(* IEC 61131-3 sources: guidance-for-physical-ai-production-designer-on-aws/source/plan2cell/examples/cell_2robot/plc/trust/head/src, 14 files *)

(* ---- E_CellError.st ---- *)
(*
 * E_CellError
 *
 * Fault codes of the cell (FB_Cell.eError), the robot drivers (FB_VassRobot.eError)
 * and the zone arbiter (FB_ZoneArbiter.eFault). ERR_NONE = no fault.
 *)

TYPE E_CellError :
(
    ERR_NONE                := 0,

    (* VASS bring-up and job handshake (FB_VassRobot) *)
    ERR_SAFETY_TIMEOUT      := 10,      (* SafeIn0.0 / SafeIn1.4 not reported *)
    ERR_DRIVES_TIMEOUT      := 11,      (* DrivesOn not reported *)
    ERR_EXT_TIMEOUT         := 12,      (* EXT mode not reported *)
    ERR_NOT_READY           := 13,      (* robot not Ready (or JobAck stuck) before a job *)
    ERR_ACK_TIMEOUT         := 14,      (* no JobAck after JobRequest *)
    ERR_ECHO_MISMATCH       := 15,      (* echoed job number <> requested job number *)
    ERR_START_TIMEOUT       := 16,      (* ProgRunning not reported after ProgStart *)
    ERR_ROBOT_STOPPED       := 17,      (* ProgRunning dropped without ProgFinished (T_STOP_DEBOUNCE) *)
    ERR_ROBOT_ERROR         := 18,      (* robot reports Error *)
    ERR_SAFETY_LOST         := 19,      (* safe status lost while up *)
    ERR_STOP_TIMEOUT        := 20,      (* robot still running after Stop + Cancel *)
    ERR_RESET_FAILED        := 21,      (* robot still in error after Reset *)
    ERR_DRIVES_LOST         := 22,      (* DrivesOn lost while up *)
    ERR_UNEXPECTED_RUN      := 23,      (* ProgRunning reported outside a job (off / bring-up / idle) *)

    (* zone protocol and supervision (FB_ZoneArbiter, FB_Cell) *)
    ERR_OP_WATCHDOG         := 30,      (* op took longer than aOps[].tLimit *)
    ERR_ZONE_WAIT_TIMEOUT   := 31,      (* zone wait past aOps[].tZoneDeadline since cycle start *)
    ERR_STEP_SEQUENCE       := 32,      (* op index did not advance by exactly +1, or 0 between two ops *)
    ERR_REQ_MISMATCH        := 33,      (* REQUEST <> mask of the reported op (debounced) *)
    ERR_TICKET_SKIPPED      := 34,      (* own ticket for another op, or zone consumed (debounced) *)
    ERR_PROGRAM_INCOMPLETE  := 35,      (* job done but last op index <> op count *)
    ERR_RELEASE_INVALID     := 36,      (* REQUEST dropped by a robot that is not running OK *)
    ERR_ROBOT_STALLED       := 37,      (* zone op without REQUEST and grant, or op index 0 too long *)
    ERR_UNEXPECTED_REQUEST  := 38,      (* holder raised bits it was not granted *)
    ERR_TICKETS_LEFT        := 39,      (* cycle done with unconsumed tickets *)
    ERR_HOME_FAILED         := 40,      (* blind homing did not reach the home pose *)
    ERR_HANDSHAKE           := 41,      (* op index changed while a grant was held (4-phase violated) *)
    ERR_ZONE_BYPASSED       := 42,      (* zone / permit op left without ever being granted *)

    (* operator *)
    ERR_OPERATOR_STOP       := 50       (* bStop *)
);
END_TYPE

(* ---- E_CellState.st ---- *)
(*
 * E_CellState
 *
 * States of the cell controller FB_Cell.
 *)

TYPE E_CellState :
(
    CS_INIT                 := 0,       (* robots off *)
    CS_BRINGUP              := 10,      (* all robots: SAFETY_ENABLE -> DRIVES_ON -> MODE_EXT -> IDLE *)
    CS_HOMING_SELECT        := 20,      (* pick robot(s) not at home *)
    CS_HOMING_RUN           := 21,      (* blind homing with HOME_FOLGE *)
    CS_READY                := 30,      (* all robots at home, waiting for start / auto-run *)
    CS_START_JOBS           := 40,      (* production Folge commanded on every active robot *)
    CS_RUNNING              := 50,      (* robots run autonomously, zones arbitrated *)
    CS_CYCLE_DONE           := 60,      (* pause T_CYCLE_PAUSE before the next cycle *)
    CS_ABORTING             := 80,      (* grants dropped, Stop + Cancel to every busy robot *)
    CS_RECOVERY             := 85,      (* after an abort mid-cycle, or a start-up with an active robot
                                           away from home: wait for bRecoveryConfirm *)
    CS_RESETTING            := 90,      (* Reset to robots in error (an operator stop cancels it) *)
    CS_ERROR                := 99       (* latched until bReset *)
);
END_TYPE

(* ---- E_GrantPolicy.st ---- *)
(*
 * E_GrantPolicy
 *
 * Zone grant policy of FB_ZoneArbiter (GVL_Cell.GRANT_POLICY).
 *)

TYPE E_GrantPolicy :
(
    GP_PLANNED  := 0,       (* zone granted only to its next ticket holder (BT order) *)
    GP_FCFS     := 1        (* oldest request first - BT order NOT enforced *)
);
END_TYPE

(* ---- E_RobotState.st ---- *)
(*
 * E_RobotState
 *
 * States of the VASS driver FB_VassRobot (one robot).
 *)

TYPE E_RobotState :
(
    RS_OFF                  := 0,       (* outputs off, waiting for bPowerOn *)
    RS_SAFETY_ENABLE        := 1,       (* SafeOut0/1 set, waiting for safe status *)
    RS_DRIVES_ON            := 2,       (* DrivesOn requested *)
    RS_MODE_EXT             := 3,       (* EXT mode requested *)
    RS_IDLE                 := 10,      (* up, no job *)
    RS_JOB_WAIT_READY       := 20,      (* waiting for Ready and no JobAck *)
    RS_JOB_SEND             := 21,      (* job number + JobRequest, waiting for JobAck *)
    RS_JOB_START            := 22,      (* ProgStart pulse *)
    RS_JOB_WAIT_RUNNING     := 23,      (* waiting for ProgRunning (or ProgFinished) *)
    RS_JOB_RUNNING          := 24,      (* program running *)
    RS_JOB_DONE             := 25,      (* ProgFinished seen, bJobDone set *)
    RS_STOPPING             := 30,      (* Stop + Cancel held *)
    RS_RESET                := 40,      (* Reset held *)
    RS_ERROR                := 99       (* latched until bCmdReset *)
);
END_TYPE

(* ---- ST_OpInfo.st ---- *)
(*
 * ST_OpInfo
 *
 * One op of one robot (GVL_Cell.aOps). Op k of robot r is
 * GVL_Cell.aOps[GVL_Cell.anRobotFirstOp[r] + k - 1].
 *)

TYPE ST_OpInfo :
STRUCT
    nRobot              : INT;      (* robot index, 1-based *)
    nOp                 : INT;      (* op index of that robot, 1-based *)
    dwZoneMask          : DWORD;    (* REQUEST/GRANT mask: zone bits 0..30, bit 31 = permit *)
    nPredFirst          : INT;      (* permit preds: GVL_Cell.aPreds[nPredFirst .. nPredFirst + nPredCount - 1] *)
    nPredCount          : INT;      (* 0 = no permit predecessors *)
    tExpected           : TIME;     (* nominal duration *)
    tLimit              : TIME;     (* op watchdog (from the grant, or from the step change if mask = 0) *)
    tZoneDeadline       : TIME;     (* latest grant time since cycle start *)
    sName               : STRING(32);
END_STRUCT
END_TYPE

(* ---- ST_RobotIn.st ---- *)
(*
 * ST_RobotIn
 *
 * Copy of one robot's input image (robot -> PLC), filled by PLC_PRG from
 * GVL_IO.bySafeIn0_<tag>..bySafeIn7_<tag> and GVL_IO.aVassInputData_<tag>.
 *)

TYPE ST_RobotIn :
STRUCT
    abySafeIn           : ARRAY[0..7] OF BYTE;      (* PROFIsafe FDIO64 safe status *)
    aVassIn             : ARRAY[0..31] OF BYTE;     (* VASS DIO256 status telegram *)
END_STRUCT
END_TYPE

(* ---- ST_RobotOut.st ---- *)
(*
 * ST_RobotOut
 *
 * One robot's output image (PLC -> robot), copied by PLC_PRG to
 * GVL_IO.bySafeOut0_<tag>..bySafeOut7_<tag> and GVL_IO.aVassOutputData_<tag>.
 *)

TYPE ST_RobotOut :
STRUCT
    abySafeOut          : ARRAY[0..7] OF BYTE;      (* PROFIsafe FDIO64 safe commands *)
    aVassOut            : ARRAY[0..31] OF BYTE;     (* VASS DIO256 command telegram *)
END_STRUCT
END_TYPE

(* ---- ST_Ticket.st ---- *)
(*
 * ST_Ticket
 *
 * One (robot, op) reference: a zone ticket in GVL_Cell.aTickets or a permit
 * predecessor in GVL_Cell.aPreds. Both indices are 1-based; 0 = none (dummy row).
 *)

TYPE ST_Ticket :
STRUCT
    nRobot              : INT;      (* robot index 1..GVL_Cell.N_ROBOTS *)
    nOp                 : INT;      (* op index of that robot 1..anRobotOpCount[nRobot] *)
END_STRUCT
END_TYPE

(* ---- GVL_Cell.st ---- *)
NAMESPACE GVL_Cell
(*
 * GVL_Cell - generated by bt2plc 0.1.0 - DO NOT EDIT
 * Plan   : bt_1791274820_cell_2robot (cell cell_2robot)
 * Grants : planned ticket order
 *)
{attribute 'qualified_only'}
VAR_GLOBAL
    (* ========================================================================
       DIMENSIONS (array bounds are literals; *_DIM >= 1)
       ======================================================================== *)
    N_ROBOTS                : INT := 1;
    N_ZONES                 : INT := 0;
    N_OPS                   : INT := 2;
    N_PREDS                 : INT := 0;

    (* ========================================================================
       PROTOCOL / TIMING
       ======================================================================== *)
    PLAN_ID                 : WORD := WORD#16#A312;             (* fold of the plan fingerprint *)
    PROD_FOLGE              : WORD := WORD#11;                  (* default production Folge *)
    HOME_FOLGE              : WORD := WORD#125;                 (* blind homing *)
    JOB_NUMBER_BYTE         : BOOL := FALSE;                    (* FALSE: WORD LE bytes 2-3, TRUE: byte 2 *)
    PROFILE_VW              : BOOL := FALSE;                    (* TRUE: VW KS24 signal map and Folge handshake instead of the simulator telegram *)
    GRANT_POLICY            : E_GrantPolicy := E_GrantPolicy#GP_PLANNED;
    HOME_SEQUENTIAL         : BOOL := TRUE;
    AUTO_RUN                : BOOL := TRUE;                     (* start the next cycle automatically *)
    STEP_BYTE               : INT := 4;                         (* robot -> PLC, WORD LE op index *)
    REQ_BYTE                : INT := 28;                        (* robot -> PLC, DWORD LE zone requests *)
    GRANT_BYTE              : INT := 12;                        (* PLC -> robot, DWORD LE zone grants *)
    PLAN_ID_BYTE            : INT := 4;                         (* PLC -> robot, WORD LE plan id *)
    PERMIT_MASK             : DWORD := DWORD#16#80000000;       (* bit 31: permit predecessors *)
    T_RESET_PULSE           : TIME := T#1S;
    T_START_PULSE           : TIME := T#500MS;
    T_STOP_PULSE            : TIME := T#1S;
    T_HANDSHAKE             : TIME := T#5S;
    T_BRINGUP_LIMIT         : TIME := T#1M;                     (* safety enable: PROFINET connection set-up *)
    T_MISMATCH_DEBOUNCE     : TIME := T#200MS;
    T_STOP_DEBOUNCE         : TIME := T#200MS;                  (* job running: ProgRunning and ProgFinished low this long = robot stopped *)
    T_CYCLE_PAUSE           : TIME := T#2S;
    T_START_LIMIT           : TIME := T#15S;
    T_ABORT_LIMIT           : TIME := T#10S;
    T_HOME_LIMIT            : TIME := T#15S500MS;

    (* ========================================================================
       VW KS24 SIGNAL INDICES (used when PROFILE_VW; $IN/$OUT index, 1-based)
       ======================================================================== *)
    VW_READY_OUT            : INT := 9;                         (* O_R_Bereit *)
    VW_RK100_OUT            : INT := 10;                        (* O_R_RK100 safety circuit *)
    VW_AUTO_OUT             : INT := 12;                        (* O_R_Auto *)
    VW_ESTOP_OUT            : INT := 13;                        (* O_R_Notaus *)
    VW_END_OUT              : INT := 14;                        (* O_R_F_ENDE / LPKT *)
    VW_PF0_OUT              : INT := 15;                        (* O_R_PFO home position *)
    VW_STEP_OUT             : INT := 97;                        (* P_PktNr_SPS op index (16 bits) *)
    VW_REL_OUT              : INT := 41;                        (* interlock releases A41-56 *)
    VW_REQ_OUT              : INT := 81;                        (* interlock requests A81-96 *)
    VW_ERR_OUT              : INT := 225;                       (* VW_FEH_BIN_A error code (8 bits) *)
    VW_DRIVES_IN            : INT := 10;                        (* I_R_Ant_Ein *)
    VW_SRB_IN               : INT := 9;                         (* I_R_SRB Folge start *)
    VW_RESET_IN             : INT := 26;                        (* I_R_Quit_St acknowledge *)
    anInterlock             : ARRAY[1..1] OF INT := [0];        (* robot r, zone z -> VW interlock 1..16 (0 = not a member): index (r-1)*1+z *)

    (* ========================================================================
       ROBOTS (index = BT order)
       ======================================================================== *)
    asRobotTag              : ARRAY[1..1] OF STRING(16) := ['R1'];
    asRobotNs               : ARRAY[1..1] OF STRING(32) := ['robot1'];
    abRobotActive           : ARRAY[1..1] OF BOOL := [TRUE];
    abSafetyBypass          : ARRAY[1..1] OF BOOL := [FALSE];   (* SIMULATION ONLY: PROFIsafe slot-1 bits not required ([[robot]] safety_bypass) *)
    awRobotProdFolge        : ARRAY[1..1] OF WORD := [WORD#11];
    anRobotFirstOp          : ARRAY[1..1] OF INT := [1];        (* op k of robot r: aOps[anRobotFirstOp[r] + k - 1] *)
    anRobotOpCount          : ARRAY[1..1] OF INT := [2];

    (* ========================================================================
       ZONES - tickets of zone z: aTickets[anZoneFirst[z] .. anZoneFirst[z] + anZoneCount[z] - 1]
       ======================================================================== *)
    asZoneName              : ARRAY[1..1] OF STRING(8) := [''];
    anZoneFirst             : ARRAY[1..1] OF INT := [0];
    anZoneCount             : ARRAY[1..1] OF INT := [0];
    aTickets                : ARRAY[1..1] OF ST_Ticket := [
        (nRobot := 0, nOp := 0)    (* no zones *)
    ];

    (* ========================================================================
       OPS - op k of robot r: aOps[anRobotFirstOp[r] + k - 1]
       ======================================================================== *)
    (* tLimit = 1.5 x tExpected + 5 s ; tZoneDeadline = 1.5 x ASAP grant + (5 + 0.2) s x depth + 10 s *)
    aOps                    : ARRAY[1..2] OF ST_OpInfo := [
        (nRobot := 1, nOp := 1, dwZoneMask := DWORD#16#00000000, nPredFirst := 0, nPredCount := 0, tExpected := T#3S729MS, tLimit := T#10S594MS, tZoneDeadline := T#10S, sName := 'STAGE_R1'),    (* R1 #1 STAGE_R1 *)
        (nRobot := 1, nOp := 2, dwZoneMask := DWORD#16#00000000, nPredFirst := 0, nPredCount := 0, tExpected := T#2S419MS, tLimit := T#8S629MS, tZoneDeadline := T#20S794MS, sName := 'HOME')    (* R1 #2 HOME *)
    ];

    (* ========================================================================
       PERMIT PREDECESSORS - op preds: aPreds[nPredFirst .. nPredFirst + nPredCount - 1]
       ======================================================================== *)
    aPreds                  : ARRAY[1..1] OF ST_Ticket := [
        (nRobot := 0, nOp := 0)    (* no permit predecessors *)
    ];
END_VAR
END_NAMESPACE

(* ---- GVL_IO.st ---- *)
NAMESPACE GVL_IO
(*
 * GVL_IO - Head PLC I/O, one block per robot
 * Generated by bt2plc 0.1.0 for cell cell_2robot (plan bt_1791274820_cell_2robot)
 *
 * This is the PROFINET Controller (master) side.
 * From the controller's perspective:
 *   "Inputs"  = data received FROM the robot device (robot status)
 *   "Outputs" = data sent TO the robot device (PLC commands)
 *
 * Map in the I/O Mapping tab of each KUKA device under the PN-Controller:
 *   SafeIO_FDIO64_<tag> inputs  -> bySafeIn0_<tag>..bySafeIn7_<tag>
 *   SafeIO_FDIO64_<tag> outputs -> bySafeOut0_<tag>..bySafeOut7_<tag>
 *   VASS_DIO256_<tag> inputs    -> aVassInputData_<tag>
 *   VASS_DIO256_<tag> outputs   -> aVassOutputData_<tag>
 *
 * Only PLC_PRG accesses this GVL: whole arrays and single bytes are copied
 * into / out of FB_Cell (never write single elements of these arrays).
 *)

{attribute 'qualified_only'}
VAR_GLOBAL

    (* ========================================================================
       R1 - robot1 - kuka_robi1 (kuka-robi1, 192.168.100.11)
       ======================================================================== *)

    (* SLOT 1 - PROFIsafe FDIO64: safe status FROM robot (8 bytes) *)
    bySafeIn0_R1            : BYTE;     (* Byte 0: Drives OK, Stopped, Reduced speed... *)
    bySafeIn1_R1            : BYTE;     (* Byte 1: Gates, E-Stop, Enabling... *)
    bySafeIn2_R1            : BYTE;     (* Byte 2: STO, SS1, SS2, SOS, SLS... *)
    bySafeIn3_R1            : BYTE;
    bySafeIn4_R1            : BYTE;
    bySafeIn5_R1            : BYTE;
    bySafeIn6_R1            : BYTE;
    bySafeIn7_R1            : BYTE;

    (* SLOT 1 - PROFIsafe FDIO64: safe commands TO robot (8 bytes) *)
    bySafeOut0_R1           : BYTE;     (* Byte 0: Drive enable, E-Stop, SS1, SS2, SLS... *)
    bySafeOut1_R1           : BYTE;     (* Byte 1: Zone enables *)
    bySafeOut2_R1           : BYTE;
    bySafeOut3_R1           : BYTE;
    bySafeOut4_R1           : BYTE;
    bySafeOut5_R1           : BYTE;
    bySafeOut6_R1           : BYTE;
    bySafeOut7_R1           : BYTE;

    (* SLOT 2 - DIO256 VASS telegram (32 bytes each direction) *)
    aVassInputData_R1       : ARRAY[0..31] OF BYTE;         (* VASS status FROM robot *)
    aVassOutputData_R1      : ARRAY[0..31] OF BYTE;         (* VASS commands TO robot *)

END_VAR
END_NAMESPACE

(* ---- FB_Cell.st ---- *)
(*
 * FB_Cell
 * Generated by bt2plc 0.1.0 for cell cell_2robot (plan bt_1791274820_cell_2robot)
 *
 * Cell control for 1 robot(s): bring-up, blind homing (HOME_FOLGE), production
 * cycle (awRobotProdFolge started on every active robot; the robots run autonomously),
 * zone / permit arbitration (FB_ZoneArbiter), supervision (op index sequence, per-op
 * watchdog, zone-wait deadline, stall, program completeness), abort (stop all, drop grants,
 * rewind tickets), recovery confirmation and reset (Reset held >= 500 ms).
 *
 *   INIT -> BRINGUP -> HOMING_SELECT <-> HOMING_RUN -> READY -> START_JOBS -> RUNNING
 *        -> CYCLE_DONE -> READY ...
 *   any fault -> ABORTING -> ERROR -(bReset)-> RESETTING -> BRINGUP -> HOMING_SELECT ...
 *   abort with a robot inside its program (op index > 0, grant held, program left
 *   incomplete or away from home), or the first bring-up after INIT (head restart /
 *   download) with an active robot away from home:
 *        ... BRINGUP -> RECOVERY -(bRecoveryConfirm)-> RESETTING -> BRINGUP -> HOMING_SELECT
 *        (operator moves the robots clear in T1 first; homing is then always sequential)
 *   Start-up homing stays automatic when every active robot is at home.
 *
 * Operator: a bStop edge is latched in every state until it is consumed - abort (normal
 * states), cancel of the reset -> ERROR (INIT / RESETTING, driver Reset low), or cleared
 * (ERROR). A bReset edge in ABORTING is applied when ERROR is reached.
 *
 * Scan order: robot drivers (commands of the previous scan) -> op index tracking ->
 * faults known so far -> arbiter (this scan's inputs, no new grants after a fault) ->
 * watchdogs -> faults -> state machine -> GRANT bytes (0 when a fault is latched).
 * Op supervision runs whenever a robot's production job is commanded / running, in any
 * cell state: op index sequence, zone ops left without grant, op index 0 while running.
 *
 * Portable: one FB_VassRobot instance per robot (no FB instance arrays), timers are
 * TIME stamps of one free-running clock (_tNow).
 *)

FUNCTION_BLOCK FB_Cell
VAR_INPUT
    bEnable             : BOOL := TRUE;
    bAutoRun            : BOOL := TRUE;     (* Level: start a cycle whenever READY *)
    bStart              : BOOL;             (* Rising edge: start one cycle *)
    bStop               : BOOL;             (* Rising edge: abort (ERR_OPERATOR_STOP) *)
    bReset              : BOOL;             (* Rising edge in CS_ERROR: reset robots and cell *)
    bRecoveryConfirm    : BOOL;             (* Rising edge (from CS_ERROR on, while bRecoveryRequired): robots cleared *)
    astIn               : ARRAY[1..1] OF ST_RobotIn;    (* Robot inputs (copied from GVL_IO) *)
END_VAR

VAR_OUTPUT
    astOut              : ARRAY[1..1] OF ST_RobotOut;   (* Robot outputs (copied to GVL_IO) *)
    eState              : E_CellState;
    eError              : E_CellError;      (* First fault, ERR_NONE when OK *)
    nErrorRobot         : INT;              (* Robot of the fault, 0 = cell *)
    nErrorOp            : INT;              (* Op index of the fault, 0 = none *)
    nErrorZone          : INT;              (* Zone of the fault, 0 = none *)
    bCycleActive        : BOOL;             (* START_JOBS or RUNNING *)
    bError              : BOOL;             (* Fault latched until the reset is done *)
    bHomingRequired     : BOOL;         (* Profile vw-ks24: a robot is not at home and must be
                                           jogged there by the operator (no blind HOME Folge) *)
    bRecoveryRequired   : BOOL;             (* bRecoveryConfirm needed before homing (abort mid-cycle / start-up away from home) *)
    udiCycles           : UDINT;            (* Completed production cycles *)
    tLastCycle          : TIME;             (* Duration of the last cycle (RUNNING) *)
    aeRobotState        : ARRAY[1..1] OF E_RobotState;
    aeRobotError        : ARRAY[1..1] OF E_CellError;
    awStep              : ARRAY[1..1] OF WORD;          (* Reported op index *)
    adwReq              : ARRAY[1..1] OF DWORD;         (* REQUEST per robot *)
    adwGrant            : ARRAY[1..1] OF DWORD;         (* GRANT per robot (as sent) *)
    anDone              : ARRAY[1..1] OF INT;           (* Ops completed in this cycle *)
    anHolder            : ARRAY[1..1] OF INT;        (* Zone holder, 0 = free *)
    anTicket            : ARRAY[1..1] OF INT;        (* Next ticket per zone *)
END_VAR

VAR
    (* ========================================================================
       ROBOT DRIVERS (one instance per robot) AND ARBITER
       ======================================================================== *)
    fbRobot_R1          : FB_VassRobot;     (* 1: robot1 - kuka_robi1 (192.168.100.11) *)
    fbArbiter           : FB_ZoneArbiter;

    (* ========================================================================
       CELL STATE
       ======================================================================== *)
    _eState             : E_CellState := E_CellState#CS_INIT;
    _eLastState         : E_CellState := E_CellState#CS_INIT;
    _bFault             : BOOL;             (* Fault latched (eError valid) *)
    _bPowerOn           : BOOL;             (* Robots: bring up *)
    _bArbReset          : BOOL := TRUE;     (* Arbiter reset in the next scan *)
    _bNeedRecovery      : BOOL;             (* Latched at an abort with a robot inside its program *)
    _bRecoveryHoming    : BOOL;             (* Homing after recovery: always sequential *)
    _bEngaged           : BOOL;             (* A robot is inside its production program / holds a grant *)
    _bConfirmLatch      : BOOL;             (* bRecoveryConfirm edge seen since CS_ERROR *)
    _bFirstBringup      : BOOL := TRUE;     (* First bring-up after CS_INIT: check the home poses *)
    _bStopReq           : BOOL;             (* bStop edge, latched until consumed *)
    _bResetReq          : BOOL;             (* bReset edge seen in CS_ABORTING, applied in CS_ERROR *)
    _bFaultScan         : BOOL;             (* Fault source known before the arbiter call (this scan) *)

    (* ========================================================================
       ROBOT STATUS (copied from the driver instances every scan)
       ======================================================================== *)
    _abIdle             : ARRAY[1..1] OF BOOL;
    _abBusy             : ARRAY[1..1] OF BOOL;
    _abDrvError         : ARRAY[1..1] OF BOOL;          (* Driver in RS_ERROR / RS_RESET *)
    _abJobActive        : ARRAY[1..1] OF BOOL;
    _abJobDone          : ARRAY[1..1] OF BOOL;
    _abAtHome           : ARRAY[1..1] OF BOOL;
    _abRobotError       : ARRAY[1..1] OF BOOL;          (* Robot reports Error *)
    _abProgRunning      : ARRAY[1..1] OF BOOL;          (* Robot reports ProgRunning *)
    _awLastStep         : ARRAY[1..1] OF WORD;

    (* ========================================================================
       COMMANDS TO THE ROBOT DRIVERS (used in the next scan)
       ======================================================================== *)
    _abJobCmd           : ARRAY[1..1] OF BOOL;
    _awJob              : ARRAY[1..1] OF WORD;
    _abProdCmd          : ARRAY[1..1] OF BOOL;          (* Commanded job is the production Folge *)
    _abStopCmd          : ARRAY[1..1] OF BOOL;
    _abResetCmd         : ARRAY[1..1] OF BOOL;
    _abHoming           : ARRAY[1..1] OF BOOL;

    (* ========================================================================
       PRODUCTION CYCLE SUPERVISION
       ======================================================================== *)
    _abHasJob           : ARRAY[1..1] OF BOOL;          (* Active robot with ops *)
    _abRobotOk          : ARRAY[1..1] OF BOOL;          (* Arbiter input *)
    _anDone             : ARRAY[1..1] OF INT;           (* Arbiter input: ops completed *)
    _anStepSeen         : ARRAY[1..1] OF INT;           (* Op index seen last scan (incl. 0) *)
    _anLastStep         : ARRAY[1..1] OF INT;           (* Last validated non-zero op index *)
    _abGranted          : ARRAY[1..1] OF BOOL;          (* Current zone op has been granted *)
    _abOpRun            : ARRAY[1..1] OF BOOL;          (* Op watchdog running *)
    _atOpStart          : ARRAY[1..1] OF TIME;
    _abStallRun         : ARRAY[1..1] OF BOOL;          (* Stall watchdog running *)
    _atStallStart       : ARRAY[1..1] OF TIME;
    _abZeroRun          : ARRAY[1..1] OF BOOL;          (* Op index 0 watchdog running *)
    _atZeroStart        : ARRAY[1..1] OF TIME;
    _tCycleStart        : TIME;

    (* ========================================================================
       TIME BASE / TIMERS / EDGES
       ======================================================================== *)
    _tonClock           : TON;              (* Free-running clock, restarted every hour *)
    _tClockBase         : TIME;
    _tNow               : TIME;             (* Monotonic time of this scan *)
    _tonState           : TON;              (* State timeout, restarts on every state change *)
    _tLimit             : TIME;
    _rtrigStart         : R_TRIG;
    _rtrigStop          : R_TRIG;
    _rtrigReset         : R_TRIG;
    _rtrigConfirm       : R_TRIG;

    (* ========================================================================
       SCRATCH
       ======================================================================== *)
    _eNew               : E_CellError;
    _nNewRobot          : INT;
    _nNewOp             : INT;
    _nHomeCount         : INT;
    _nDone              : INT;
    _r                  : INT;
    _iOp                : INT;
    _nStep              : INT;
    _nPrev              : INT;              (* Op index that is left *)
    _tZeroLimit         : TIME;
    _dwGrant            : DWORD;
    _bBypass            : BOOL;
    _bAll               : BOOL;
    _bSequential        : BOOL;

    (* Profile vw-ks24: interlock grant / partner release encoding *)
    _z                  : INT;
    _q                  : INT;
    _nIl                : INT;
    _nIlQ               : INT;
    _nIdx               : INT;
    _nB                 : INT;
    _nBit               : INT;
    _wBits              : WORD;
    _bGrantBit          : BOOL;
    _bPartner           : BOOL;
END_VAR
(*
 * FB_Cell - Implementation
 *)

IF NOT bEnable THEN
    _eState := E_CellState#CS_INIT;
END_IF

(* ============================================================================
   TIME BASE / EDGES
   ============================================================================ *)
_tonClock(IN := TRUE, PT := T#1H);
_tNow := _tClockBase + _tonClock.ET;
IF _tonClock.Q THEN
    _tClockBase := _tNow;
    _tonClock(IN := FALSE);
    _tonClock(IN := TRUE, PT := T#1H);
END_IF

_rtrigStart(CLK := bStart);
_rtrigStop(CLK := bStop);
_rtrigReset(CLK := bReset);
_rtrigConfirm(CLK := bRecoveryConfirm);

(* Operator stop: latched in every state until consumed (abort, cancelled reset, CS_ERROR);
   it also cancels a reset that is pending from CS_ABORTING *)
IF _rtrigStop.Q THEN
    _bStopReq := TRUE;
    _bResetReq := FALSE;
END_IF

FOR _r := 1 TO GVL_Cell.N_ROBOTS DO
    _abHasJob[_r] := GVL_Cell.abRobotActive[_r] AND (GVL_Cell.anRobotOpCount[_r] > 0);
END_FOR

(* ============================================================================
   ROBOT DRIVERS (commands from the previous scan; GRANT bytes are added below)
   ============================================================================ *)

(* 1: R1 - robot1 *)
fbRobot_R1(
    bEnable     := bEnable,
    bPowerOn    := _bPowerOn,
    bCmdJob     := _abJobCmd[1],
    wJobNr      := _awJob[1],
    bProdJob    := _abProdCmd[1],
    bCmdStop    := _abStopCmd[1],
    bCmdReset   := _abResetCmd[1],
    nRobot      := 1,
    stIn        := astIn[1]);
astOut[1]         := fbRobot_R1.stOut;
aeRobotState[1]   := fbRobot_R1.eState;
aeRobotError[1]   := fbRobot_R1.eError;
awStep[1]         := fbRobot_R1.wStep;
adwReq[1]         := fbRobot_R1.dwZoneReq;
_awLastStep[1]    := fbRobot_R1.wLastStep;
_abIdle[1]        := fbRobot_R1.bIdle;
_abBusy[1]        := fbRobot_R1.bBusy;
_abDrvError[1]    := fbRobot_R1.bError;
_abJobActive[1]   := fbRobot_R1.bJobActive;
_abJobDone[1]     := fbRobot_R1.bJobDone;
_abAtHome[1]      := fbRobot_R1.bAtHome;
_abRobotError[1]  := fbRobot_R1.bRobotError;
_abProgRunning[1] := fbRobot_R1.bProgRunning;

(* A robot inside its production program or holding a grant (previous scan's commands):
   inside an op, between two ops, finished with an incomplete program, or left the
   home pose during the current cycle *)
_bEngaged := FALSE;
FOR _r := 1 TO GVL_Cell.N_ROBOTS DO
    IF _abJobCmd[_r] AND _abProdCmd[_r] THEN
        IF awStep[_r] <> WORD#0 THEN
            _bEngaged := TRUE;
        ELSIF (_awLastStep[_r] <> WORD#0) AND NOT _abJobDone[_r] THEN
            _bEngaged := TRUE;
        ELSIF _abJobDone[_r] AND (WORD_TO_INT(_awLastStep[_r]) <> GVL_Cell.anRobotOpCount[_r]) THEN
            _bEngaged := TRUE;
        ELSIF NOT _abAtHome[_r]
              AND ((_awLastStep[_r] <> WORD#0) OR (_anLastStep[_r] <> 0) OR _abJobActive[_r]) THEN
            _bEngaged := TRUE;
        END_IF
    END_IF
    IF fbArbiter.adwGrant[_r] <> DWORD#0 THEN
        _bEngaged := TRUE;
    END_IF
END_FOR

(* ============================================================================
   OP INDEX TRACKING (production job commanded, any cell state)
   The index must advance by exactly +1. The op that is left (also at the job end,
   index -> 0) must have been granted if it has a zone / permit mask (both policies).
   Index 0 while the program runs is valid only before the first / after the last op.
   ============================================================================ *)
_eNew := E_CellError#ERR_NONE;
_nNewRobot := 0;
_nNewOp := 0;
FOR _r := 1 TO GVL_Cell.N_ROBOTS DO
    IF _abJobCmd[_r] AND _abProdCmd[_r] THEN
        _nStep := WORD_TO_INT(awStep[_r]);
        IF _nStep <> _anStepSeen[_r] THEN
            _nPrev := _anStepSeen[_r];
            _bBypass := FALSE;
            IF (_nPrev >= 1) AND (_nPrev <= GVL_Cell.anRobotOpCount[_r]) AND NOT _abGranted[_r] THEN
                _iOp := GVL_Cell.anRobotFirstOp[_r] + _nPrev - 1;
                IF GVL_Cell.aOps[_iOp].dwZoneMask <> DWORD#0 THEN
                    _bBypass := TRUE;               (* zone / permit op left without a grant *)
                END_IF
            END_IF
            IF _bBypass THEN
                IF _eNew = E_CellError#ERR_NONE THEN
                    _eNew := E_CellError#ERR_ZONE_BYPASSED;
                    _nNewRobot := _r;
                    _nNewOp := _nPrev;
                END_IF
            ELSIF _nStep <> 0 THEN
                IF (_nStep = _anLastStep[_r] + 1) AND (_nStep <= GVL_Cell.anRobotOpCount[_r]) THEN
                    _anLastStep[_r] := _nStep;
                ELSIF _eNew = E_CellError#ERR_NONE THEN
                    _eNew := E_CellError#ERR_STEP_SEQUENCE;
                    _nNewRobot := _r;
                    _nNewOp := _nStep;
                END_IF
            END_IF
            _anStepSeen[_r] := _nStep;
            _abGranted[_r] := FALSE;
            _abOpRun[_r] := FALSE;
            _abStallRun[_r] := FALSE;
            _abZeroRun[_r] := FALSE;
        END_IF

        (* index 0 while the program runs, between two ops *)
        IF _abJobActive[_r] AND (_nStep = 0) AND (_anLastStep[_r] > 0)
           AND (_anLastStep[_r] < GVL_Cell.anRobotOpCount[_r])
           AND (_eNew = E_CellError#ERR_NONE) THEN
            _eNew := E_CellError#ERR_STEP_SEQUENCE;
            _nNewRobot := _r;
            _nNewOp := 0;
        END_IF

        (* ops completed (permit predecessors): validated index - 1, all at job done *)
        IF _abJobDone[_r] AND (_anLastStep[_r] = GVL_Cell.anRobotOpCount[_r]) THEN
            _nDone := GVL_Cell.anRobotOpCount[_r];
        ELSIF _anLastStep[_r] > 0 THEN
            _nDone := _anLastStep[_r] - 1;
        ELSE
            _nDone := 0;
        END_IF
        _anDone[_r] := MAX(_anDone[_r], _nDone);
    END_IF
END_FOR

(* ============================================================================
   ZONE ARBITER (this scan's robot inputs)
   No new grants in a scan in which the cell already knows it will abort:
   driver error, latched operator stop, latched fault, supervision fault above.
   ============================================================================ *)
_bFaultScan := _bFault OR _bStopReq OR (_eNew <> E_CellError#ERR_NONE);
FOR _r := 1 TO GVL_Cell.N_ROBOTS DO
    _abRobotOk[_r] := _abJobActive[_r] AND _abJobCmd[_r] AND _abProdCmd[_r] AND NOT _abRobotError[_r];
    IF _abDrvError[_r] THEN
        _bFaultScan := TRUE;
    END_IF
END_FOR
fbArbiter(
    bReset      := _bArbReset,
    bEnable     := ((_eState = E_CellState#CS_START_JOBS) OR (_eState = E_CellState#CS_RUNNING))
                   AND NOT _bFaultScan,
    ePolicy     := GVL_Cell.GRANT_POLICY,
    tDebounce   := GVL_Cell.T_MISMATCH_DEBOUNCE,
    tNow        := _tNow,
    abRobotOk   := _abRobotOk,
    awStep      := awStep,
    adwReq      := adwReq,
    anDone      := _anDone);
_bArbReset := FALSE;

(* ============================================================================
   WATCHDOGS (production job running, any cell state)
   op watchdog from the step change (mask 0) or from the grant; stall; zone wait;
   op index 0: T_HANDSHAKE before the first op, MAX(last op tLimit, T_HANDSHAKE)
   after the last op
   ============================================================================ *)
FOR _r := 1 TO GVL_Cell.N_ROBOTS DO
    IF _abJobCmd[_r] AND _abProdCmd[_r] AND _abJobActive[_r] THEN
        _nStep := _anStepSeen[_r];
        IF (_nStep >= 1) AND (_nStep <= GVL_Cell.anRobotOpCount[_r]) THEN
            _iOp := GVL_Cell.anRobotFirstOp[_r] + _nStep - 1;
            IF GVL_Cell.aOps[_iOp].dwZoneMask = DWORD#0 THEN
                IF NOT _abOpRun[_r] THEN
                    _abOpRun[_r] := TRUE;
                    _atOpStart[_r] := _tNow;
                END_IF
            ELSE
                IF fbArbiter.adwGrant[_r] <> DWORD#0 THEN
                    _abGranted[_r] := TRUE;
                END_IF
                IF _abGranted[_r] AND NOT _abOpRun[_r] THEN
                    _abOpRun[_r] := TRUE;
                    _atOpStart[_r] := _tNow;
                END_IF

                (* zone op with neither REQUEST nor grant *)
                IF NOT _abGranted[_r] AND (adwReq[_r] = DWORD#0) THEN
                    IF NOT _abStallRun[_r] THEN
                        _abStallRun[_r] := TRUE;
                        _atStallStart[_r] := _tNow;
                    ELSIF ((_tNow - _atStallStart[_r]) >= GVL_Cell.T_HANDSHAKE)
                          AND (_eNew = E_CellError#ERR_NONE) THEN
                        _eNew := E_CellError#ERR_ROBOT_STALLED;
                        _nNewRobot := _r;
                        _nNewOp := _nStep;
                    END_IF
                ELSE
                    _abStallRun[_r] := FALSE;
                END_IF

                (* zone wait past the deadline (measured since the cycle started RUNNING) *)
                IF NOT _abGranted[_r] AND (adwReq[_r] <> DWORD#0)
                   AND (_eState = E_CellState#CS_RUNNING)
                   AND ((_tNow - _tCycleStart) > GVL_Cell.aOps[_iOp].tZoneDeadline)
                   AND (_eNew = E_CellError#ERR_NONE) THEN
                    _eNew := E_CellError#ERR_ZONE_WAIT_TIMEOUT;
                    _nNewRobot := _r;
                    _nNewOp := _nStep;
                END_IF
            END_IF

            IF _abOpRun[_r] AND ((_tNow - _atOpStart[_r]) >= GVL_Cell.aOps[_iOp].tLimit)
               AND (_eNew = E_CellError#ERR_NONE) THEN
                _eNew := E_CellError#ERR_OP_WATCHDOG;
                _nNewRobot := _r;
                _nNewOp := _nStep;
            END_IF
        ELSIF _nStep = 0 THEN
            (* program running without an op: before the first / after the last op *)
            IF NOT _abZeroRun[_r] THEN
                _abZeroRun[_r] := TRUE;
                _atZeroStart[_r] := _tNow;
            END_IF
            _tZeroLimit := GVL_Cell.T_HANDSHAKE;
            IF (_anLastStep[_r] >= 1) AND (_anLastStep[_r] = GVL_Cell.anRobotOpCount[_r]) THEN
                _iOp := GVL_Cell.anRobotFirstOp[_r] + _anLastStep[_r] - 1;
                IF GVL_Cell.aOps[_iOp].tLimit > _tZeroLimit THEN
                    _tZeroLimit := GVL_Cell.aOps[_iOp].tLimit;
                END_IF
            END_IF
            IF ((_tNow - _atZeroStart[_r]) >= _tZeroLimit) AND (_eNew = E_CellError#ERR_NONE) THEN
                _eNew := E_CellError#ERR_ROBOT_STALLED;
                _nNewRobot := _r;
                _nNewOp := 0;
            END_IF
        END_IF
    ELSE
        _abZeroRun[_r] := FALSE;
    END_IF
END_FOR

(* ============================================================================
   FAULT COLLECTION (first wins: robot > supervision > arbiter > operator)
   ============================================================================ *)
IF (_eState <> E_CellState#CS_INIT) AND (_eState <> E_CellState#CS_ABORTING)
   AND (_eState <> E_CellState#CS_ERROR) AND (_eState <> E_CellState#CS_RESETTING) THEN
    FOR _r := 1 TO GVL_Cell.N_ROBOTS DO
        IF _abDrvError[_r] AND NOT _bFault AND (_eState <> E_CellState#CS_RECOVERY) THEN
            _bFault := TRUE;
            eError := aeRobotError[_r];
            nErrorRobot := _r;
            nErrorOp := WORD_TO_INT(awStep[_r]);
            nErrorZone := 0;
        END_IF
    END_FOR
    IF (_eNew <> E_CellError#ERR_NONE) AND NOT _bFault THEN
        _bFault := TRUE;
        eError := _eNew;
        nErrorRobot := _nNewRobot;
        nErrorOp := _nNewOp;
        nErrorZone := 0;
    END_IF
    IF fbArbiter.bFault AND NOT _bFault THEN
        _bFault := TRUE;
        eError := fbArbiter.eFault;
        nErrorRobot := fbArbiter.nFaultRobot;
        nErrorOp := 0;
        IF (fbArbiter.nFaultRobot >= 1) AND (fbArbiter.nFaultRobot <= GVL_Cell.N_ROBOTS) THEN
            nErrorOp := WORD_TO_INT(awStep[fbArbiter.nFaultRobot]);
        END_IF
        nErrorZone := fbArbiter.nFaultZone;
    END_IF
    IF _bStopReq THEN
        _bStopReq := FALSE;                 (* consumed by this abort *)
        IF NOT _bFault THEN
            _bFault := TRUE;
            eError := E_CellError#ERR_OPERATOR_STOP;
            nErrorRobot := 0;
            nErrorOp := 0;
            nErrorZone := 0;
        END_IF
    END_IF
    IF _bFault THEN
        _eState := E_CellState#CS_ABORTING;
    END_IF
END_IF

(* ============================================================================
   STATE TIMER (after the transitions above: a new state starts with a fresh timer)
   ============================================================================ *)
IF _eState <> _eLastState THEN
    IF _eState = E_CellState#CS_ABORTING THEN
        _bConfirmLatch := FALSE;
        IF _bEngaged THEN
            _bNeedRecovery := TRUE;         (* aborted with a robot inside its program *)
        END_IF
    END_IF
    _tonState(IN := FALSE);
    _eLastState := _eState;
END_IF
CASE _eState OF
E_CellState#CS_HOMING_RUN:
    _tLimit := GVL_Cell.T_HOME_LIMIT;
E_CellState#CS_START_JOBS:
    _tLimit := GVL_Cell.T_START_LIMIT;
E_CellState#CS_CYCLE_DONE:
    _tLimit := GVL_Cell.T_CYCLE_PAUSE;
E_CellState#CS_ABORTING, E_CellState#CS_RESETTING:
    _tLimit := GVL_Cell.T_ABORT_LIMIT;
ELSE
    _tLimit := T#24H;
END_CASE
_tonState(IN := TRUE, PT := _tLimit);

(* Recovery confirm: accepted once the robots are stopped (CS_ERROR on), used in CS_RECOVERY *)
IF _rtrigConfirm.Q AND _bNeedRecovery
   AND ((_eState = E_CellState#CS_ERROR) OR (_eState = E_CellState#CS_RESETTING)
        OR (_eState = E_CellState#CS_BRINGUP) OR (_eState = E_CellState#CS_RECOVERY)) THEN
    _bConfirmLatch := TRUE;
END_IF

(* ============================================================================
   STATE MACHINE
   ============================================================================ *)
CASE _eState OF

E_CellState#CS_INIT:
    _bPowerOn := FALSE;
    _bArbReset := TRUE;
    _bFirstBringup := TRUE;                 (* head start / restart: robot poses unknown *)
    FOR _r := 1 TO GVL_Cell.N_ROBOTS DO
        _abJobCmd[_r] := FALSE;
        _abProdCmd[_r] := FALSE;
        _abStopCmd[_r] := FALSE;
        _abResetCmd[_r] := FALSE;
        _abHoming[_r] := FALSE;
    END_FOR
    IF bEnable THEN
        IF _bStopReq THEN
            (* operator stop before the start-up: no automatic bring-up *)
            _bStopReq := FALSE;
            _bResetReq := FALSE;
            _bFault := TRUE;
            eError := E_CellError#ERR_OPERATOR_STOP;
            nErrorRobot := 0;
            nErrorOp := 0;
            nErrorZone := 0;
            _eState := E_CellState#CS_ERROR;
        ELSE
            _eState := E_CellState#CS_BRINGUP;
        END_IF
    END_IF

E_CellState#CS_BRINGUP:
    _bPowerOn := TRUE;
    _bAll := TRUE;
    FOR _r := 1 TO GVL_Cell.N_ROBOTS DO
        IF NOT _abIdle[_r] THEN
            _bAll := FALSE;
        END_IF
    END_FOR
    IF _bAll THEN
        IF _bFirstBringup THEN
            (* first bring-up after INIT: any robot away from home (also an idle one)
               may stand anywhere in the shared space (head restart / download mid-cycle) *)
            _bFirstBringup := FALSE;
            FOR _r := 1 TO GVL_Cell.N_ROBOTS DO
                IF NOT _abAtHome[_r] AND NOT _bNeedRecovery THEN
                    _bNeedRecovery := TRUE;
                    _bConfirmLatch := FALSE;
                END_IF
            END_FOR
        END_IF
        IF _bNeedRecovery THEN
            _eState := E_CellState#CS_RECOVERY;
        ELSE
            _eState := E_CellState#CS_HOMING_SELECT;
        END_IF
    END_IF

E_CellState#CS_RECOVERY:
    (* robots may be anywhere inside the shared space: the operator moves them
       clear (T1, driver errors are ignored here) and confirms; then the drivers
       are reset, brought up again and blind homing runs one robot at a time *)
    IF _bConfirmLatch THEN
        _bConfirmLatch := FALSE;
        _bNeedRecovery := FALSE;
        _bRecoveryHoming := TRUE;
        _eState := E_CellState#CS_RESETTING;
    END_IF

E_CellState#CS_HOMING_SELECT:
    IF GVL_Cell.PROFILE_VW THEN
        (* VW cell.src starts a Folge only once the robot reports PF0, and there is no blind
           home Folge: wait for the operator to jog every robot home (ERR_HOME_FAILED on
           T_HOME_LIMIT tells which robot is not at home). *)
        _bAll := TRUE;
        FOR _r := 1 TO GVL_Cell.N_ROBOTS DO
            IF NOT _abAtHome[_r] THEN
                _bAll := FALSE;
                bHomingRequired := TRUE;
            END_IF
        END_FOR
        IF _bAll THEN
            bHomingRequired := FALSE;
            _bRecoveryHoming := FALSE;
            _eState := E_CellState#CS_READY;
        ELSIF _tonState.Q THEN
            _bFault := TRUE;
            eError := E_CellError#ERR_HOME_FAILED;
            nErrorRobot := 0;
            FOR _r := GVL_Cell.N_ROBOTS TO 1 BY -1 DO
                IF NOT _abAtHome[_r] THEN
                    nErrorRobot := _r;
                END_IF
            END_FOR
            nErrorOp := 0;
            nErrorZone := 0;
            _eState := E_CellState#CS_ERROR;
        END_IF
    ELSE
        _bSequential := GVL_Cell.HOME_SEQUENTIAL OR _bRecoveryHoming;
        _nHomeCount := 0;
        FOR _r := 1 TO GVL_Cell.N_ROBOTS DO
            _abHoming[_r] := FALSE;
            IF NOT _abAtHome[_r] AND (NOT _bSequential OR (_nHomeCount = 0)) THEN
                _abHoming[_r] := TRUE;
                _awJob[_r] := GVL_Cell.HOME_FOLGE;
                _abProdCmd[_r] := FALSE;
                _nHomeCount := _nHomeCount + 1;
            END_IF
        END_FOR
        IF _nHomeCount = 0 THEN
            _bRecoveryHoming := FALSE;
            _eState := E_CellState#CS_READY;
        ELSE
            _eState := E_CellState#CS_HOMING_RUN;
        END_IF
    END_IF

E_CellState#CS_HOMING_RUN:
    _bAll := TRUE;
    FOR _r := 1 TO GVL_Cell.N_ROBOTS DO
        IF _abHoming[_r] THEN
            _abJobCmd[_r] := TRUE;
            IF NOT _abJobDone[_r] THEN
                _bAll := FALSE;
            ELSIF NOT _abAtHome[_r] AND NOT _bFault THEN
                _bFault := TRUE;
                eError := E_CellError#ERR_HOME_FAILED;
                nErrorRobot := _r;
                nErrorOp := 0;
                nErrorZone := 0;
            END_IF
        END_IF
    END_FOR
    IF _bFault THEN
        _eState := E_CellState#CS_ABORTING;
    ELSIF _bAll THEN
        FOR _r := 1 TO GVL_Cell.N_ROBOTS DO
            IF _abHoming[_r] THEN
                _abJobCmd[_r] := FALSE;
                _abHoming[_r] := FALSE;
            END_IF
        END_FOR
        _eState := E_CellState#CS_HOMING_SELECT;
    ELSIF _tonState.Q THEN
        _bFault := TRUE;
        eError := E_CellError#ERR_HOME_FAILED;
        nErrorRobot := 0;
        FOR _r := GVL_Cell.N_ROBOTS TO 1 BY -1 DO
            IF _abHoming[_r] AND NOT _abJobDone[_r] THEN
                nErrorRobot := _r;
            END_IF
        END_FOR
        nErrorOp := 0;
        nErrorZone := 0;
        _eState := E_CellState#CS_ABORTING;
    END_IF

E_CellState#CS_READY:
    IF _rtrigStart.Q OR bAutoRun THEN
        _bAll := TRUE;
        FOR _r := 1 TO GVL_Cell.N_ROBOTS DO
            IF _abHasJob[_r] AND NOT _abAtHome[_r] THEN
                _bAll := FALSE;             (* programs start at the home pose *)
            END_IF
        END_FOR
        IF _bAll THEN
            _bArbReset := TRUE;             (* rewind tickets for this cycle *)
            FOR _r := 1 TO GVL_Cell.N_ROBOTS DO
                _anStepSeen[_r] := 0;
                _anLastStep[_r] := 0;
                _anDone[_r] := 0;
                _abGranted[_r] := FALSE;
                _abOpRun[_r] := FALSE;
                _abStallRun[_r] := FALSE;
                _abZeroRun[_r] := FALSE;
                _abProdCmd[_r] := FALSE;
                IF _abHasJob[_r] THEN
                    _awJob[_r] := GVL_Cell.awRobotProdFolge[_r];
                    _abProdCmd[_r] := TRUE;
                END_IF
            END_FOR
            _eState := E_CellState#CS_START_JOBS;
        ELSE
            _eState := E_CellState#CS_HOMING_SELECT;
        END_IF
    END_IF

E_CellState#CS_START_JOBS:
    _bAll := TRUE;
    FOR _r := 1 TO GVL_Cell.N_ROBOTS DO
        IF _abHasJob[_r] THEN
            _abJobCmd[_r] := TRUE;
            IF NOT (_abJobActive[_r] OR _abJobDone[_r]) THEN
                _bAll := FALSE;
            END_IF
        END_IF
    END_FOR
    IF _bAll THEN
        _tCycleStart := _tNow;
        _eState := E_CellState#CS_RUNNING;
    ELSIF _tonState.Q THEN
        _bFault := TRUE;
        eError := E_CellError#ERR_START_TIMEOUT;
        nErrorRobot := 0;
        FOR _r := GVL_Cell.N_ROBOTS TO 1 BY -1 DO
            IF _abHasJob[_r] AND NOT (_abJobActive[_r] OR _abJobDone[_r]) THEN
                nErrorRobot := _r;
            END_IF
        END_FOR
        nErrorOp := 0;
        nErrorZone := 0;
        _eState := E_CellState#CS_ABORTING;
    END_IF

E_CellState#CS_RUNNING:
    _bAll := TRUE;
    FOR _r := 1 TO GVL_Cell.N_ROBOTS DO
        IF _abHasJob[_r] THEN
            IF NOT _abJobDone[_r] THEN
                _bAll := FALSE;
            ELSIF (WORD_TO_INT(_awLastStep[_r]) <> GVL_Cell.anRobotOpCount[_r]) AND NOT _bFault THEN
                _bFault := TRUE;
                eError := E_CellError#ERR_PROGRAM_INCOMPLETE;
                nErrorRobot := _r;
                nErrorOp := WORD_TO_INT(_awLastStep[_r]);
                nErrorZone := 0;
            END_IF
        END_IF
    END_FOR
    IF _bFault THEN
        _eState := E_CellState#CS_ABORTING;
    ELSIF _bAll THEN
        IF NOT fbArbiter.bAllConsumed THEN
            _bFault := TRUE;
            eError := E_CellError#ERR_TICKETS_LEFT;
            nErrorRobot := 0;
            nErrorOp := 0;
            nErrorZone := 0;
            _eState := E_CellState#CS_ABORTING;
        ELSE
            FOR _r := 1 TO GVL_Cell.N_ROBOTS DO
                _abJobCmd[_r] := FALSE;
            END_FOR
            udiCycles := udiCycles + 1;
            tLastCycle := _tNow - _tCycleStart;
            _eState := E_CellState#CS_CYCLE_DONE;
        END_IF
    END_IF

E_CellState#CS_CYCLE_DONE:
    IF _tonState.Q THEN
        _eState := E_CellState#CS_READY;
    END_IF

E_CellState#CS_ABORTING:
    _bArbReset := TRUE;                     (* drop all grants, rewind tickets *)
    _bAll := TRUE;
    FOR _r := 1 TO GVL_Cell.N_ROBOTS DO
        _abJobCmd[_r] := FALSE;
        _abHoming[_r] := FALSE;
        _abStopCmd[_r] := TRUE;
        IF _abBusy[_r] THEN
            _bAll := FALSE;
        END_IF
    END_FOR
    IF _rtrigReset.Q AND NOT _rtrigStop.Q THEN
        _bResetReq := TRUE;                 (* applied once CS_ERROR is reached *)
        _bStopReq := FALSE;                 (* the abort in progress already stops *)
    END_IF
    IF _bAll OR _tonState.Q THEN
        _eState := E_CellState#CS_ERROR;
    END_IF

E_CellState#CS_ERROR:
    _bArbReset := TRUE;
    FOR _r := 1 TO GVL_Cell.N_ROBOTS DO
        _abStopCmd[_r] := FALSE;            (* drivers keep Stop while a robot still runs *)
        _abResetCmd[_r] := FALSE;           (* re-arm the reset edges *)
    END_FOR
    IF _bStopReq THEN
        _bStopReq := FALSE;                 (* already stopped *)
        _bResetReq := FALSE;
    ELSIF _rtrigReset.Q OR _bResetReq THEN
        _bResetReq := FALSE;
        _eState := E_CellState#CS_RESETTING;
    END_IF

E_CellState#CS_RESETTING:
    IF _bStopReq THEN
        (* operator stop cancels the reset: driver Reset low, no bring-up / homing *)
        _bStopReq := FALSE;
        _bResetReq := FALSE;
        FOR _r := 1 TO GVL_Cell.N_ROBOTS DO
            _abResetCmd[_r] := FALSE;
        END_FOR
        IF _bRecoveryHoming THEN
            _bRecoveryHoming := FALSE;
            _bNeedRecovery := TRUE;         (* confirm again after the next reset *)
        END_IF
        _bConfirmLatch := FALSE;
        _bFault := TRUE;
        eError := E_CellError#ERR_OPERATOR_STOP;
        nErrorRobot := 0;
        nErrorOp := 0;
        nErrorZone := 0;
        _eState := E_CellState#CS_ERROR;
    ELSE
        _bAll := TRUE;
        FOR _r := 1 TO GVL_Cell.N_ROBOTS DO
            _abResetCmd[_r] := _abDrvError[_r];
            IF _abDrvError[_r] OR _abBusy[_r] OR _abProgRunning[_r] THEN
                _bAll := FALSE;
            END_IF
        END_FOR
        IF _bAll THEN
            FOR _r := 1 TO GVL_Cell.N_ROBOTS DO
                _abResetCmd[_r] := FALSE;
                _abProdCmd[_r] := FALSE;
            END_FOR
            _bFault := FALSE;
            eError := E_CellError#ERR_NONE;
            nErrorRobot := 0;
            nErrorOp := 0;
            nErrorZone := 0;
            _bArbReset := TRUE;
            _eState := E_CellState#CS_BRINGUP;  (* then recovery (if needed) or blind homing *)
        ELSIF _tonState.Q THEN
            IF NOT _bFault THEN                 (* reset after a recovery confirm failed *)
                _bFault := TRUE;
                eError := E_CellError#ERR_RESET_FAILED;
                nErrorRobot := 0;
                FOR _r := GVL_Cell.N_ROBOTS TO 1 BY -1 DO
                    IF _abDrvError[_r] OR _abBusy[_r] OR _abProgRunning[_r] THEN
                        nErrorRobot := _r;
                    END_IF
                END_FOR
                nErrorOp := 0;
                nErrorZone := 0;
            END_IF
            _eState := E_CellState#CS_ERROR;
        END_IF
    END_IF

END_CASE

(* ============================================================================
   GRANT BYTES (PLC -> robot, DWORD LE): non-zero only while the job runs and no
   fault is latched (also covers faults decided after the arbiter in this scan)
   ============================================================================ *)
FOR _r := 1 TO GVL_Cell.N_ROBOTS DO
    IF _abJobActive[_r] AND NOT _bFault AND NOT _bFaultScan THEN
        _dwGrant := fbArbiter.adwGrant[_r];
    ELSE
        _dwGrant := DWORD#0;
    END_IF
    adwGrant[_r] := _dwGrant;
    IF GVL_Cell.PROFILE_VW THEN
        (* Per interlock n of robot r: grant E(80+n) = the arbiter's zone bit, partner release
           E(40+n) = AND of the releases A(40+n) of the other members of that zone (the robot
           waits for it before it enters, and its online driving condition keeps watching it). *)
        FOR _z := 1 TO GVL_Cell.N_ZONES DO
            _nIl := GVL_Cell.anInterlock[(_r - 1) * GVL_Cell.N_ZONES + _z];
            IF (_nIl >= 1) AND (_nIl <= 16) THEN
                _bGrantBit := (_dwGrant AND SHL(DWORD#1, _z - 1)) <> DWORD#0;
                _bPartner := TRUE;
                FOR _q := 1 TO GVL_Cell.N_ROBOTS DO
                    IF _q <> _r THEN
                        _nIlQ := GVL_Cell.anInterlock[(_q - 1) * GVL_Cell.N_ZONES + _z];
                        IF (_nIlQ >= 1) AND (_nIlQ <= 16) THEN
                            _nIdx := GVL_Cell.VW_REL_OUT + _nIlQ - 1;
                            _nB := (_nIdx - 1) / 8;
                            _nBit := (_nIdx - 1) MOD 8;
                            IF (SHR(BYTE_TO_WORD(astIn[_q].aVassIn[_nB]), _nBit) AND WORD#1) = WORD#0 THEN
                                _bPartner := FALSE;
                            END_IF
                        END_IF
                    END_IF
                END_FOR
                _nIdx := GVL_Cell.VW_REQ_OUT + _nIl - 1;
                _nB := (_nIdx - 1) / 8;
                _nBit := (_nIdx - 1) MOD 8;
                IF _bGrantBit THEN
                    _wBits := BYTE_TO_WORD(astOut[_r].aVassOut[_nB]) OR SHL(WORD#1, _nBit);
                    astOut[_r].aVassOut[_nB] := WORD_TO_BYTE(_wBits);
                END_IF
                _nIdx := GVL_Cell.VW_REL_OUT + _nIl - 1;
                _nB := (_nIdx - 1) / 8;
                _nBit := (_nIdx - 1) MOD 8;
                IF _bPartner AND NOT _bFault AND NOT _bFaultScan THEN
                    _wBits := BYTE_TO_WORD(astOut[_r].aVassOut[_nB]) OR SHL(WORD#1, _nBit);
                    astOut[_r].aVassOut[_nB] := WORD_TO_BYTE(_wBits);
                END_IF
            END_IF
        END_FOR
    ELSE
        astOut[_r].aVassOut[GVL_Cell.GRANT_BYTE]     := DWORD_TO_BYTE(_dwGrant AND DWORD#16#FF);
        astOut[_r].aVassOut[GVL_Cell.GRANT_BYTE + 1] := DWORD_TO_BYTE(SHR(_dwGrant, 8) AND DWORD#16#FF);
        astOut[_r].aVassOut[GVL_Cell.GRANT_BYTE + 2] := DWORD_TO_BYTE(SHR(_dwGrant, 16) AND DWORD#16#FF);
        astOut[_r].aVassOut[GVL_Cell.GRANT_BYTE + 3] := DWORD_TO_BYTE(SHR(_dwGrant, 24) AND DWORD#16#FF);
    END_IF
END_FOR

(* ============================================================================
   OUTPUTS
   ============================================================================ *)
eState := _eState;
bError := _bFault;
bCycleActive := (_eState = E_CellState#CS_START_JOBS) OR (_eState = E_CellState#CS_RUNNING);
bRecoveryRequired := _bNeedRecovery;
anHolder := fbArbiter.anHolder;
anTicket := fbArbiter.anTicket;
anDone := _anDone;
END_FUNCTION_BLOCK

(* ---- FB_VassRobot.st ---- *)
(*
 * FB_VassRobot
 * Generated by bt2plc 0.1.0 for cell cell_2robot (plan bt_1791274820_cell_2robot)
 *
 * VW VASS protocol driver for ONE robot (KUKA VKRC nexxt V8.2 DIM 2 via PROFINET).
 * Portable: no pointers, no REFERENCE, no OOP - the robot IO is passed as struct
 * copies (stIn / stOut) by the caller (FB_Cell, PLC_PRG copies GVL_IO).
 *
 *   Bring-up : SAFETY_ENABLE (T_BRINGUP_LIMIT: PROFINET / PROFIsafe connection set-up)
 *              -> DRIVES_ON -> MODE_EXT -> IDLE   (T_HANDSHAKE each)
 *   Job      : WAIT_READY -> SEND (echo checked) -> START (T_START_PULSE) -> WAIT_RUNNING
 *              -> RUNNING -> DONE   (WAIT_RUNNING -> DONE if the job finished between scans)
 *              (RUNNING -> ERROR ERR_ROBOT_STOPPED only after ProgRunning and ProgFinished
 *              stayed low for T_STOP_DEBOUNCE: a robot may publish the two bits in different
 *              bus frames at the Folge end)
 *              (T_HANDSHAKE per handshake state)
 *   Abort    : STOPPING (Stop + Cancel held >= T_STOP_PULSE and until ProgRunning drops)
 *   Recovery : ERROR -> RESET (Reset held T_RESET_PULSE >= 500 ms while bCmdReset stays TRUE;
 *              bCmdReset dropped = reset cancelled -> ERROR) -> SAFETY_ENABLE
 *              (still ProgRunning after the pulse -> ERROR, ERR_STOP_TIMEOUT)
 *   Command handshake: bCmdJob is a level request (rising edge latched),
 *              bJobDone the acknowledge (cleared while bCmdJob = FALSE).
 *
 * Stop is never dropped while the robot still reports ProgRunning (also in ERROR / RESET).
 * ProgRunning outside a job (OFF, bring-up, IDLE) -> ERROR (ERR_UNEXPECTED_RUN, Stop + Cancel).
 * The zone GRANT bytes (GVL_Cell.GRANT_BYTE .. +3) are written 0 here: FB_Cell encodes
 * them after FB_ZoneArbiter has run, so a grant reaches the robot in the scan it is computed.
 *
 * Profile vw-ks24 (GVL_Cell.PROFILE_VW): the VW tech package on the robot does the Folge
 * handshake, so the signal map and the job states differ (same state names):
 *   status  : ready A9, safety A10 + A13, auto A12, home A15 (PF0), Folge end A14,
 *             echo PRG_NR_REFL A1-8, op index P_PktNr_SPS, error code VW_FEH_BIN_A
 *   commands: drives E10, Folge number PRG_NR E1-8, start SRB E9 (level), reset E26
 *   job     : SEND writes PRG_NR and waits for the echo; START holds SRB until the robot
 *             leaves home (its cycle-start point clears PF0); RUNNING waits for Folge end;
 *             DONE clears PRG_NR and waits for the Folge end to fall
 *   zones   : REQUEST bit z is synthesised as "requesting or occupying",
 *             A(80+n) OR NOT A(40+n), which is exactly the REQUEST semantics of the arbiter;
 *             the release is A(40+n) going TRUE again. There is no 4-phase handshake.
 *   stop    : no Stop/Cancel bits exist; the head drops the drives, withdraws the partner
 *             releases (the robot's online driving condition stops it on the path) and clears
 *             PRG_NR. Recovery needs manual homing (PF0), there is no blind HOME Folge.
 *)

FUNCTION_BLOCK FB_VassRobot
VAR_INPUT
    bEnable             : BOOL := TRUE;
    nRobot              : INT := 1;         (* 1-based robot index (profile vw-ks24: interlock map) *)
    bPowerOn            : BOOL;             (* Level: bring the robot up *)
    bCmdJob             : BOOL;             (* Level request (rising edge latched): run job wJobNr *)
    wJobNr              : WORD;             (* Folge number, latched at job accept *)
    bProdJob            : BOOL;             (* wJobNr is the production Folge: send PLAN_ID, track wLastStep *)
    bCmdStop            : BOOL;             (* Level: abort the active job *)
    bCmdReset           : BOOL;             (* Rising edge in RS_ERROR: reset the robot; hold until bError drops *)
    stIn                : ST_RobotIn;       (* Copy of this robot's GVL_IO inputs *)
END_VAR

VAR_OUTPUT
    stOut               : ST_RobotOut;      (* Copy to this robot's GVL_IO outputs (GRANT bytes = 0) *)
    eState              : E_RobotState;
    eError              : E_CellError;
    bIdle               : BOOL;
    bBusy               : BOOL;             (* Job, stopping or resetting *)
    bJobActive          : BOOL;             (* Job started and ProgRunning *)
    bJobDone            : BOOL;             (* Job finished (cleared while bCmdJob = FALSE) *)
    bError              : BOOL;             (* RS_ERROR or RS_RESET *)

    (* Decoded robot status *)
    bDrivesOn           : BOOL;
    bProgRunning        : BOOL;
    bAtHome             : BOOL;
    bModeExt            : BOOL;
    bRobotReady         : BOOL;
    bRobotError         : BOOL;
    bProgFinished       : BOOL;
    bJobAck             : BOOL;
    bSafetyOK           : BOOL;
    wActiveJob          : WORD;             (* Echoed job number *)
    wStep               : WORD;             (* Reported op index, 0 = no program *)
    wLastStep           : WORD;             (* Max op index of the running production job (cleared at job accept) *)
    dwZoneReq           : DWORD;            (* REQUEST DWORD: zone bits 0..30, permit bit 31 *)
    wRobotErrorCode     : WORD;
END_VAR

VAR
    _eState             : E_RobotState := E_RobotState#RS_OFF;
    _eLastState         : E_RobotState := E_RobotState#RS_OFF;
    _wJob               : WORD;             (* Job number latched at accept *)
    _bProdJob           : BOOL;             (* Latched bProdJob *)
    _bJobPending        : BOOL;             (* Job edge seen, not yet accepted *)
    _bInJob             : BOOL;
    _bUp                : BOOL;
    _bNoJob             : BOOL;             (* Off / bring-up / idle: ProgRunning is not expected *)

    (* Commands to the robot *)
    _bSafeEnable        : BOOL;
    _bDrivesOnCmd       : BOOL;
    _bExtCmd            : BOOL;
    _bStartCmd          : BOOL;
    _bStopCmd           : BOOL;
    _bCancelCmd         : BOOL;
    _bResetCmd          : BOOL;
    _bJobReqCmd         : BOOL;

    (* Timers *)
    _tonStep            : TON;              (* State timeout, restarts on every state change *)
    _tonPulse           : TON;              (* Start / stop / reset pulse width *)
    _tonStopDebounce    : TON;              (* RS_JOB_RUNNING: ProgRunning + ProgFinished low (T_STOP_DEBOUNCE) *)
    _tStepLimit         : TIME;

    (* Edge detection *)
    _rtrigJob           : R_TRIG;
    _rtrigReset         : R_TRIG;

    (* Profile vw-ks24 *)
    _bFolgeEnd          : BOOL;             (* A14 Folge end *)
    _bVwStarted         : BOOL;             (* SRB acknowledged: the robot left its home point *)
    _nIdx               : INT;              (* signal index 1..256 *)
    _nB                 : INT;              (* telegram byte of _nIdx *)
    _nBit               : INT;              (* bit of _nIdx *)
    _wTmp               : WORD;
    _bTmp               : BOOL;
    _z                  : INT;
    _n                  : INT;

    _i                  : INT;
END_VAR
(*
 * FB_VassRobot - Implementation
 * Reads the robot status from stIn, writes the commands to stOut.
 *)

IF NOT bEnable THEN
    FOR _i := 0 TO 31 DO
        stOut.aVassOut[_i] := BYTE#0;
    END_FOR
    FOR _i := 0 TO 7 DO
        stOut.abySafeOut[_i] := BYTE#0;
    END_FOR
    _eState := E_RobotState#RS_OFF;
    _eLastState := E_RobotState#RS_OFF;
    _bJobPending := FALSE;
    eState := _eState;
    eError := E_CellError#ERR_NONE;
    bIdle := FALSE;
    bBusy := FALSE;
    bJobActive := FALSE;
    bJobDone := FALSE;
    bError := FALSE;
    wLastStep := WORD#0;
    RETURN;
END_IF

(* ============================================================================
   DECODE ROBOT STATUS (robot -> PLC)
   ============================================================================ *)

(* The job state of the scan we start in (the global transitions below may change it); the
   vw-ks24 decode needs it for the "occupied" term. *)
_bInJob := (_eState = E_RobotState#RS_JOB_WAIT_READY) OR (_eState = E_RobotState#RS_JOB_SEND)
           OR (_eState = E_RobotState#RS_JOB_START) OR (_eState = E_RobotState#RS_JOB_WAIT_RUNNING)
           OR (_eState = E_RobotState#RS_JOB_RUNNING);

IF GVL_Cell.PROFILE_VW THEN
    (* ---- VW KS24 signal map (status bits addressed by $OUT index) ---- *)
    _nIdx := GVL_Cell.VW_READY_OUT;
    _nB := (_nIdx - 1) / 8;
    _nBit := (_nIdx - 1) MOD 8;
    bRobotReady := (SHR(BYTE_TO_WORD(stIn.aVassIn[_nB]), _nBit) AND WORD#1) = WORD#1;

    _nIdx := GVL_Cell.VW_AUTO_OUT;
    _nB := (_nIdx - 1) / 8;
    _nBit := (_nIdx - 1) MOD 8;
    bModeExt := (SHR(BYTE_TO_WORD(stIn.aVassIn[_nB]), _nBit) AND WORD#1) = WORD#1;

    _nIdx := GVL_Cell.VW_PF0_OUT;
    _nB := (_nIdx - 1) / 8;
    _nBit := (_nIdx - 1) MOD 8;
    bAtHome := (SHR(BYTE_TO_WORD(stIn.aVassIn[_nB]), _nBit) AND WORD#1) = WORD#1;

    _nIdx := GVL_Cell.VW_END_OUT;
    _nB := (_nIdx - 1) / 8;
    _nBit := (_nIdx - 1) MOD 8;
    _bFolgeEnd := (SHR(BYTE_TO_WORD(stIn.aVassIn[_nB]), _nBit) AND WORD#1) = WORD#1;
    bProgFinished := _bFolgeEnd;

    (* A10 (RK100: user_saf and em_stop group) is the drive / safety-circuit feedback; A9
       (Bereit) drops while a Folge runs, so it is only used for the job handshake. *)
    _nIdx := GVL_Cell.VW_RK100_OUT;
    _nB := (_nIdx - 1) / 8;
    _nBit := (_nIdx - 1) MOD 8;
    _bTmp := (SHR(BYTE_TO_WORD(stIn.aVassIn[_nB]), _nBit) AND WORD#1) = WORD#1;
    bDrivesOn := _bTmp;
    _nIdx := GVL_Cell.VW_ESTOP_OUT;
    _nB := (_nIdx - 1) / 8;
    _nBit := (_nIdx - 1) MOD 8;
    bSafetyOK := _bTmp AND ((SHR(BYTE_TO_WORD(stIn.aVassIn[_nB]), _nBit) AND WORD#1) = WORD#1)
                 AND stIn.abySafeIn[0].0 AND stIn.abySafeIn[1].4;

    (* Echo: PRG_NR_REFL A1-8 *)
    wActiveJob := BYTE_TO_WORD(stIn.aVassIn[0]);
    bJobAck := (wActiveJob <> WORD#0) AND (wActiveJob = _wJob);

    (* Op index: P_PktNr_SPS, 16 bits little-endian from VW_STEP_OUT *)
    _nB := (GVL_Cell.VW_STEP_OUT - 1) / 8;
    wStep := BYTE_TO_WORD(stIn.aVassIn[_nB]) OR SHL(BYTE_TO_WORD(stIn.aVassIn[_nB + 1]), 8);

    (* Error code: VW_FEH_BIN_A, 8 bits *)
    _nB := (GVL_Cell.VW_ERR_OUT - 1) / 8;
    wRobotErrorCode := BYTE_TO_WORD(stIn.aVassIn[_nB]);
    bRobotError := wRobotErrorCode <> WORD#0;

    (* REQUEST bit z = A(80+n) OR NOT A(40+n): requesting, or inside ("occupied"). The
       release is A(40+n) going TRUE again, which drops the bit. The "occupied" term counts
       only while this driver has a job: an all-zero frame (robot not connected yet, PROFINET
       down) would otherwise read as "inside every interlock". *)
    dwZoneReq := DWORD#0;
    FOR _z := 1 TO GVL_Cell.N_ZONES DO
        _n := GVL_Cell.anInterlock[(nRobot - 1) * GVL_Cell.N_ZONES + _z];
        IF (_n >= 1) AND (_n <= 16) THEN
            _nIdx := GVL_Cell.VW_REQ_OUT + _n - 1;
            _nB := (_nIdx - 1) / 8;
            _nBit := (_nIdx - 1) MOD 8;
            _bTmp := (SHR(BYTE_TO_WORD(stIn.aVassIn[_nB]), _nBit) AND WORD#1) = WORD#1;
            _nIdx := GVL_Cell.VW_REL_OUT + _n - 1;
            _nB := (_nIdx - 1) / 8;
            _nBit := (_nIdx - 1) MOD 8;
            IF _bTmp OR (_bInJob AND ((SHR(BYTE_TO_WORD(stIn.aVassIn[_nB]), _nBit) AND WORD#1) = WORD#0)) THEN
                dwZoneReq := dwZoneReq OR SHL(DWORD#1, _z - 1);
            END_IF
        END_IF
    END_FOR

    (* No ProgRunning bit: the Folge runs while its number is echoed and the robot is neither
       at its home point nor reporting the Folge end. *)
    bProgRunning := (wActiveJob <> WORD#0) AND (wActiveJob = _wJob) AND NOT bAtHome
                    AND NOT _bFolgeEnd;
ELSE
    (* Status word byte 0 / 1 *)
    bDrivesOn     := stIn.aVassIn[0].0;
    bProgRunning  := stIn.aVassIn[0].1;
    bAtHome       := stIn.aVassIn[0].2;
    bModeExt      := stIn.aVassIn[0].4;
    bRobotReady   := stIn.aVassIn[0].5;
    bRobotError   := stIn.aVassIn[0].6;
    bProgFinished := stIn.aVassIn[1].2;
    bJobAck       := stIn.aVassIn[1].3;

    (* Echoed job number from bytes 2-3 (or byte 2 only) *)
    IF GVL_Cell.JOB_NUMBER_BYTE THEN
        wActiveJob := BYTE_TO_WORD(stIn.aVassIn[2]);
    ELSE
        wActiveJob := BYTE_TO_WORD(stIn.aVassIn[2])
                      OR SHL(BYTE_TO_WORD(stIn.aVassIn[3]), 8);
    END_IF

    (* Op index (WORD LE) and zone REQUEST (DWORD LE) *)
    wStep := BYTE_TO_WORD(stIn.aVassIn[GVL_Cell.STEP_BYTE])
             OR SHL(BYTE_TO_WORD(stIn.aVassIn[GVL_Cell.STEP_BYTE + 1]), 8);

    dwZoneReq := BYTE_TO_DWORD(stIn.aVassIn[GVL_Cell.REQ_BYTE])
                 OR SHL(BYTE_TO_DWORD(stIn.aVassIn[GVL_Cell.REQ_BYTE + 1]), 8)
                 OR SHL(BYTE_TO_DWORD(stIn.aVassIn[GVL_Cell.REQ_BYTE + 2]), 16)
                 OR SHL(BYTE_TO_DWORD(stIn.aVassIn[GVL_Cell.REQ_BYTE + 3]), 24);

    (* Error code from bytes 10-11 *)
    wRobotErrorCode := BYTE_TO_WORD(stIn.aVassIn[10])
                       OR SHL(BYTE_TO_WORD(stIn.aVassIn[11]), 8);

    (* Safety status: SafeIn0.0 drives OK, SafeIn1.4 E-Stop OK *)
    bSafetyOK := stIn.abySafeIn[0].0 AND stIn.abySafeIn[1].4;
END_IF

(* SIMULATION ONLY (bt2plc [[robot]] safety_bypass -> GVL_Cell.abSafetyBypass, e.g. a KUKA virtual controller whose FDIO64
   slot carries no F-data to this non-safety controller): the slot-1 bits are not required. The
   vw-ks24 drive / E-stop status bits still count. *)
IF (nRobot >= 1) AND (nRobot <= GVL_Cell.N_ROBOTS) AND GVL_Cell.abSafetyBypass[nRobot] THEN
    IF GVL_Cell.PROFILE_VW THEN
        _nIdx := GVL_Cell.VW_ESTOP_OUT;
        _nB := (_nIdx - 1) / 8;
        _nBit := (_nIdx - 1) MOD 8;
        bSafetyOK := bDrivesOn AND ((SHR(BYTE_TO_WORD(stIn.aVassIn[_nB]), _nBit) AND WORD#1) = WORD#1);
    ELSE
        bSafetyOK := TRUE;
    END_IF
END_IF

(* ============================================================================
   EDGES
   ============================================================================ *)
_rtrigJob(CLK := bCmdJob);
_rtrigReset(CLK := bCmdReset);
IF _rtrigJob.Q THEN
    _bJobPending := TRUE;
END_IF
IF NOT bCmdJob THEN
    _bJobPending := FALSE;
END_IF

(* ============================================================================
   GLOBAL TRANSITIONS
   ============================================================================ *)
_bInJob := (_eState = E_RobotState#RS_JOB_WAIT_READY) OR (_eState = E_RobotState#RS_JOB_SEND)
           OR (_eState = E_RobotState#RS_JOB_START) OR (_eState = E_RobotState#RS_JOB_WAIT_RUNNING)
           OR (_eState = E_RobotState#RS_JOB_RUNNING);
_bUp := _bInJob OR (_eState = E_RobotState#RS_IDLE);
_bNoJob := (_eState = E_RobotState#RS_OFF) OR (_eState = E_RobotState#RS_SAFETY_ENABLE)
           OR (_eState = E_RobotState#RS_DRIVES_ON) OR (_eState = E_RobotState#RS_MODE_EXT)
           OR (_eState = E_RobotState#RS_IDLE);

IF _bInJob AND bCmdStop THEN
    _eState := E_RobotState#RS_STOPPING;
ELSIF _bUp AND bRobotError THEN
    eError := E_CellError#ERR_ROBOT_ERROR;
    _eState := E_RobotState#RS_ERROR;
ELSIF _bUp AND NOT bSafetyOK THEN
    eError := E_CellError#ERR_SAFETY_LOST;
    _eState := E_RobotState#RS_ERROR;
ELSIF _bUp AND NOT bDrivesOn THEN
    eError := E_CellError#ERR_DRIVES_LOST;
    _eState := E_RobotState#RS_ERROR;
ELSIF _bNoJob AND bProgRunning AND NOT GVL_Cell.PROFILE_VW THEN
    (* a program runs that this driver did not start (head restart / download, manual
       start): RS_ERROR holds Stop + Cancel while ProgRunning *)
    eError := E_CellError#ERR_UNEXPECTED_RUN;
    _eState := E_RobotState#RS_ERROR;
END_IF

(* ============================================================================
   STATE TIMER (after the global transitions: a new state always starts with
   fresh timers, also when it was entered by a global transition this scan)
   ============================================================================ *)
IF _eState <> _eLastState THEN
    _tonStep(IN := FALSE);
    _tonPulse(IN := FALSE);
    _tonStopDebounce(IN := FALSE);
    _eLastState := _eState;
END_IF
IF _eState = E_RobotState#RS_STOPPING THEN
    _tStepLimit := GVL_Cell.T_ABORT_LIMIT;
ELSIF _eState = E_RobotState#RS_SAFETY_ENABLE THEN
    _tStepLimit := GVL_Cell.T_BRINGUP_LIMIT;    (* PROFINET / PROFIsafe connection set-up *)
ELSE
    _tStepLimit := GVL_Cell.T_HANDSHAKE;        (* drives / EXT and job handshakes *)
END_IF
_tonStep(IN := TRUE, PT := _tStepLimit);

(* ============================================================================
   STATE MACHINE
   ============================================================================ *)
CASE _eState OF

E_RobotState#RS_OFF:
    _bSafeEnable := FALSE;
    _bDrivesOnCmd := FALSE;
    _bExtCmd := FALSE;
    _bJobReqCmd := FALSE;
    _bStartCmd := FALSE;
    _bStopCmd := FALSE;
    _bCancelCmd := FALSE;
    _bResetCmd := FALSE;
    IF bPowerOn THEN
        _eState := E_RobotState#RS_SAFETY_ENABLE;
    END_IF

E_RobotState#RS_SAFETY_ENABLE:
    _bSafeEnable := TRUE;
    IF bSafetyOK THEN
        _eState := E_RobotState#RS_DRIVES_ON;
    ELSIF _tonStep.Q THEN
        eError := E_CellError#ERR_SAFETY_TIMEOUT;
        _eState := E_RobotState#RS_ERROR;
    END_IF

E_RobotState#RS_DRIVES_ON:
    _bDrivesOnCmd := TRUE;
    IF bDrivesOn THEN
        _eState := E_RobotState#RS_MODE_EXT;
    ELSIF _tonStep.Q THEN
        eError := E_CellError#ERR_DRIVES_TIMEOUT;
        _eState := E_RobotState#RS_ERROR;
    END_IF

E_RobotState#RS_MODE_EXT:
    _bExtCmd := TRUE;
    IF bModeExt THEN
        _eState := E_RobotState#RS_IDLE;
    ELSIF _tonStep.Q THEN
        eError := E_CellError#ERR_EXT_TIMEOUT;
        _eState := E_RobotState#RS_ERROR;
    END_IF

E_RobotState#RS_IDLE:
    _bJobReqCmd := FALSE;
    _bStartCmd := FALSE;
    _bStopCmd := FALSE;
    _bCancelCmd := FALSE;
    IF NOT bCmdJob THEN
        bJobDone := FALSE;
    END_IF
    IF NOT bPowerOn THEN
        _eState := E_RobotState#RS_OFF;
    ELSIF _bJobPending THEN
        _bJobPending := FALSE;
        _wJob := wJobNr;
        _bProdJob := bProdJob;
        bJobDone := FALSE;
        wLastStep := WORD#0;
        _eState := E_RobotState#RS_JOB_WAIT_READY;
    END_IF

E_RobotState#RS_JOB_WAIT_READY:
    _bJobReqCmd := FALSE;                   (* guarantees a rising edge in RS_JOB_SEND *)
    _bVwStarted := FALSE;
    IF GVL_Cell.PROFILE_VW THEN
        (* the robot waits at its home point with PRG_NR_REFL = 0 *)
        IF bRobotReady AND bAtHome AND (wActiveJob = WORD#0) THEN
            _eState := E_RobotState#RS_JOB_SEND;
        ELSIF _tonStep.Q THEN
            eError := E_CellError#ERR_NOT_READY;
            _eState := E_RobotState#RS_ERROR;
        END_IF
    ELSIF bRobotReady AND NOT bJobAck THEN
        _eState := E_RobotState#RS_JOB_SEND;
    ELSIF _tonStep.Q THEN
        eError := E_CellError#ERR_NOT_READY;
        _eState := E_RobotState#RS_ERROR;
    END_IF

E_RobotState#RS_JOB_SEND:
    _bJobReqCmd := TRUE;                    (* vw: PRG_NR is written in the encode section *)
    IF GVL_Cell.PROFILE_VW THEN
        (* the robot mirrors PRG_NR on A1-8 while it waits for the Folge start *)
        IF wActiveJob = _wJob THEN
            _eState := E_RobotState#RS_JOB_START;
        ELSIF _tonStep.Q THEN
            eError := E_CellError#ERR_ACK_TIMEOUT;
            _eState := E_RobotState#RS_ERROR;
        END_IF
    ELSIF bJobAck THEN
        _bJobReqCmd := FALSE;
        IF wActiveJob = _wJob THEN
            _eState := E_RobotState#RS_JOB_START;
        ELSE
            eError := E_CellError#ERR_ECHO_MISMATCH;
            _eState := E_RobotState#RS_ERROR;
        END_IF
    ELSIF _tonStep.Q THEN
        _bJobReqCmd := FALSE;
        eError := E_CellError#ERR_ACK_TIMEOUT;
        _eState := E_RobotState#RS_ERROR;
    END_IF

E_RobotState#RS_JOB_START:
    _bStartCmd := TRUE;
    IF GVL_Cell.PROFILE_VW THEN
        (* SRB stays a level until the robot leaves its home point (its cycle start clears PF0) *)
        _bJobReqCmd := TRUE;                (* keep PRG_NR *)
        IF NOT bAtHome THEN
            _bVwStarted := TRUE;
            _bStartCmd := FALSE;
            _eState := E_RobotState#RS_JOB_RUNNING;
        ELSIF _tonStep.Q THEN
            eError := E_CellError#ERR_START_TIMEOUT;
            _eState := E_RobotState#RS_ERROR;
        END_IF
    ELSE
        _bJobReqCmd := FALSE;
        _tonPulse(IN := TRUE, PT := GVL_Cell.T_START_PULSE);
        IF _tonPulse.Q THEN
            _bStartCmd := FALSE;
            _eState := E_RobotState#RS_JOB_WAIT_RUNNING;
        END_IF
    END_IF

E_RobotState#RS_JOB_WAIT_RUNNING:
    _bStartCmd := FALSE;
    IF bProgRunning THEN
        _eState := E_RobotState#RS_JOB_RUNNING;
    ELSIF bProgFinished THEN
        (* finished between two scans - the robot clears ProgFinished on job accept *)
        _eState := E_RobotState#RS_JOB_DONE;
    ELSIF _tonStep.Q THEN
        eError := E_CellError#ERR_START_TIMEOUT;
        _eState := E_RobotState#RS_ERROR;
    END_IF

E_RobotState#RS_JOB_RUNNING:
    (* no timeout here: per-op watchdogs in FB_Cell, HOME uses T_HOME_LIMIT *)
    IF GVL_Cell.PROFILE_VW THEN
        _bJobReqCmd := TRUE;                (* keep PRG_NR until the Folge end *)
        IF _bFolgeEnd THEN
            _eState := E_RobotState#RS_JOB_DONE;
        END_IF
    ELSE
        (* ProgRunning low without ProgFinished is a stop only when it lasts T_STOP_DEBOUNCE:
           the robot writes the two bits to its outputs one after the other (KRL submit), so a
           bus frame taken between them shows both low for one cycle at a normal Folge end. *)
        _tonStopDebounce(IN := NOT bProgRunning AND NOT bProgFinished, PT := GVL_Cell.T_STOP_DEBOUNCE);
        IF bProgFinished AND NOT bProgRunning THEN
            _eState := E_RobotState#RS_JOB_DONE;
        ELSIF _tonStopDebounce.Q THEN
            eError := E_CellError#ERR_ROBOT_STOPPED;
            _eState := E_RobotState#RS_ERROR;
        END_IF
    END_IF

E_RobotState#RS_JOB_DONE:
    IF GVL_Cell.PROFILE_VW THEN
        (* clear PRG_NR, then wait for the Folge end (A14) to fall before the next job *)
        _bJobReqCmd := FALSE;
        IF NOT _bFolgeEnd THEN
            bJobDone := TRUE;
            _eState := E_RobotState#RS_IDLE;
        ELSIF _tonStep.Q THEN
            eError := E_CellError#ERR_HANDSHAKE;
            _eState := E_RobotState#RS_ERROR;
        END_IF
    ELSE
        bJobDone := TRUE;
        _eState := E_RobotState#RS_IDLE;
    END_IF

E_RobotState#RS_STOPPING:
    _bJobReqCmd := FALSE;                   (* vw: clears PRG_NR; FB_Cell withdraws the grants
                                               and partner releases, which stops the robot on
                                               its path through its own driving condition *)
    _bStartCmd := FALSE;
    _bStopCmd := TRUE;
    _bCancelCmd := TRUE;
    IF GVL_Cell.PROFILE_VW THEN
        _bDrivesOnCmd := FALSE;             (* no Stop/Cancel bits in KS24: drop the drives *)
    END_IF
    _tonPulse(IN := TRUE, PT := GVL_Cell.T_STOP_PULSE);
    IF _tonPulse.Q AND NOT bProgRunning THEN
        _bStopCmd := FALSE;
        _bCancelCmd := FALSE;
        _eState := E_RobotState#RS_IDLE;
    ELSIF _tonStep.Q THEN
        (* keep Stop + Cancel: RS_ERROR holds them while ProgRunning *)
        eError := E_CellError#ERR_STOP_TIMEOUT;
        _eState := E_RobotState#RS_ERROR;
    END_IF

E_RobotState#RS_ERROR:
    _bJobReqCmd := FALSE;
    _bStartCmd := FALSE;
    _bStopCmd := bProgRunning;              (* never drop Stop while the robot still runs *)
    _bCancelCmd := bProgRunning;
    _bResetCmd := FALSE;
    IF _rtrigReset.Q THEN
        _eState := E_RobotState#RS_RESET;
    END_IF

E_RobotState#RS_RESET:
    _bStopCmd := bProgRunning;
    _bCancelCmd := bProgRunning;
    (* DrivesOn low while Reset is held: a KUKA controller switches the drives on only at a rising edge of
       $DRIVES_ON after the messages are acknowledged ($CONF_MESS), so RS_DRIVES_ON must raise it again *)
    _bDrivesOnCmd := FALSE;
    _bResetCmd := TRUE;                     (* held >= 500 ms - robot requirement *)
    _tonPulse(IN := TRUE, PT := GVL_Cell.T_RESET_PULSE);
    IF NOT bCmdReset THEN
        (* reset withdrawn by the cell (operator stop): Reset low, error kept *)
        _bResetCmd := FALSE;
        _eState := E_RobotState#RS_ERROR;
    ELSIF _tonPulse.Q THEN
        _bResetCmd := FALSE;
        IF bProgRunning THEN
            (* never leave the error with a running program: RS_ERROR keeps Stop + Cancel *)
            eError := E_CellError#ERR_STOP_TIMEOUT;
            _eState := E_RobotState#RS_ERROR;
        ELSIF NOT bRobotError THEN
            eError := E_CellError#ERR_NONE;
            _eState := E_RobotState#RS_SAFETY_ENABLE;
        ELSE
            eError := E_CellError#ERR_RESET_FAILED;
            _eState := E_RobotState#RS_ERROR;
        END_IF
    END_IF

END_CASE

(* ============================================================================
   JOB STATUS
   ============================================================================ *)
_bInJob := (_eState = E_RobotState#RS_JOB_WAIT_READY) OR (_eState = E_RobotState#RS_JOB_SEND)
           OR (_eState = E_RobotState#RS_JOB_START) OR (_eState = E_RobotState#RS_JOB_WAIT_RUNNING)
           OR (_eState = E_RobotState#RS_JOB_RUNNING);
bJobActive := bProgRunning AND ((_eState = E_RobotState#RS_JOB_START)
              OR (_eState = E_RobotState#RS_JOB_WAIT_RUNNING) OR (_eState = E_RobotState#RS_JOB_RUNNING));

(* Latched max op index of the running production job (step 0 = between jobs) *)
IF bJobActive AND _bProdJob AND (wStep > wLastStep) THEN
    wLastStep := wStep;
END_IF

(* ============================================================================
   ENCODE COMMANDS (PLC -> robot)
   ============================================================================ *)
IF GVL_Cell.PROFILE_VW THEN
    (* ---- VW KS24 commands: PRG_NR A1-8, SRB, drives, acknowledge ---- *)
    FOR _i := 0 TO 31 DO
        stOut.aVassOut[_i] := BYTE#0;
    END_FOR
    (* PRG_NR only from RS_JOB_SEND on: in RS_JOB_WAIT_READY the robot must still echo 0
       (it picks the number up through cell.src as soon as it is written). *)
    IF _bJobReqCmd THEN
        stOut.aVassOut[0] := WORD_TO_BYTE(_wJob AND WORD#16#FF);
    END_IF
    _nIdx := GVL_Cell.VW_SRB_IN;
    _nB := (_nIdx - 1) / 8;
    _nBit := (_nIdx - 1) MOD 8;
    IF _bStartCmd THEN
        _wTmp := BYTE_TO_WORD(stOut.aVassOut[_nB]) OR SHL(WORD#1, _nBit);
        stOut.aVassOut[_nB] := WORD_TO_BYTE(_wTmp);
    END_IF
    _nIdx := GVL_Cell.VW_DRIVES_IN;
    _nB := (_nIdx - 1) / 8;
    _nBit := (_nIdx - 1) MOD 8;
    IF _bDrivesOnCmd THEN
        _wTmp := BYTE_TO_WORD(stOut.aVassOut[_nB]) OR SHL(WORD#1, _nBit);
        stOut.aVassOut[_nB] := WORD_TO_BYTE(_wTmp);
    END_IF
    _nIdx := GVL_Cell.VW_RESET_IN;
    _nB := (_nIdx - 1) / 8;
    _nBit := (_nIdx - 1) MOD 8;
    IF _bResetCmd THEN
        _wTmp := BYTE_TO_WORD(stOut.aVassOut[_nB]) OR SHL(WORD#1, _nBit);
        stOut.aVassOut[_nB] := WORD_TO_BYTE(_wTmp);
    END_IF
    (* PLAN_ID on a free telegram byte pair, only with the production job (0 = no check) *)
    IF (GVL_Cell.PLAN_ID_BYTE > 0) AND _bInJob AND _bProdJob THEN
        stOut.aVassOut[GVL_Cell.PLAN_ID_BYTE]     := WORD_TO_BYTE(GVL_Cell.PLAN_ID AND WORD#16#FF);
        stOut.aVassOut[GVL_Cell.PLAN_ID_BYTE + 1] := WORD_TO_BYTE(SHR(GVL_Cell.PLAN_ID, 8) AND WORD#16#FF);
    END_IF
    (* The interlock grants E(80+n) and partner releases E(40+n) are written by FB_Cell. *)
ELSE
stOut.aVassOut[0].0 := _bDrivesOnCmd;
stOut.aVassOut[0].1 := _bStartCmd;
stOut.aVassOut[0].2 := _bStopCmd;
stOut.aVassOut[0].3 := _bCancelCmd;
stOut.aVassOut[0].4 := _bExtCmd;
stOut.aVassOut[0].5 := _bResetCmd;
stOut.aVassOut[0].6 := FALSE;               (* homing uses HOME_FOLGE, not HomeRequest *)
(* MoveEnable: held in every state but RS_OFF, also through a reset (DrivesOn drops there for the
   $DRIVES_ON edge). A KUKA KSS 9.2 maps $MOVE_ENABLE to it: it refuses EXT with $MOVE_ENABLE on the
   always-TRUE $IN[1025] (M_249), and a motion enable that dropped with DrivesOn needs a new
   acknowledgement (M_1210) before the drives come on. The robot simulator ignores this bit. *)
stOut.aVassOut[0].7 := _eState <> E_RobotState#RS_OFF;
stOut.aVassOut[1].0 := _bJobReqCmd;

(* Job number, bytes 2-3 (or byte 2 only) *)
IF _bInJob THEN
    stOut.aVassOut[2] := WORD_TO_BYTE(_wJob AND WORD#16#FF);
    IF GVL_Cell.JOB_NUMBER_BYTE THEN
        stOut.aVassOut[3] := BYTE#0;
    ELSE
        stOut.aVassOut[3] := WORD_TO_BYTE(SHR(_wJob, 8) AND WORD#16#FF);
    END_IF
ELSE
    stOut.aVassOut[2] := BYTE#0;
    stOut.aVassOut[3] := BYTE#0;
END_IF

(* PLAN_ID, only with the production job *)
IF _bInJob AND _bProdJob THEN
    stOut.aVassOut[GVL_Cell.PLAN_ID_BYTE]     := WORD_TO_BYTE(GVL_Cell.PLAN_ID AND WORD#16#FF);
    stOut.aVassOut[GVL_Cell.PLAN_ID_BYTE + 1] := WORD_TO_BYTE(SHR(GVL_Cell.PLAN_ID, 8) AND WORD#16#FF);
ELSE
    stOut.aVassOut[GVL_Cell.PLAN_ID_BYTE]     := BYTE#0;
    stOut.aVassOut[GVL_Cell.PLAN_ID_BYTE + 1] := BYTE#0;
END_IF

(* GRANT bytes: encoded by FB_Cell after FB_ZoneArbiter *)
stOut.aVassOut[GVL_Cell.GRANT_BYTE]     := BYTE#0;
stOut.aVassOut[GVL_Cell.GRANT_BYTE + 1] := BYTE#0;
stOut.aVassOut[GVL_Cell.GRANT_BYTE + 2] := BYTE#0;
stOut.aVassOut[GVL_Cell.GRANT_BYTE + 3] := BYTE#0;
END_IF

(* Safe outputs *)
IF _bSafeEnable THEN
    stOut.abySafeOut[0] := BYTE#16#01;      (* drive enable *)
    stOut.abySafeOut[1] := BYTE#16#0F;      (* zones 1-4 enable *)
ELSE
    stOut.abySafeOut[0] := BYTE#0;
    stOut.abySafeOut[1] := BYTE#0;
END_IF

(* ============================================================================
   PUBLISH
   ============================================================================ *)
eState := _eState;
bIdle  := (_eState = E_RobotState#RS_IDLE);
bBusy  := _bInJob OR (_eState = E_RobotState#RS_STOPPING) OR (_eState = E_RobotState#RS_RESET);
bError := (_eState = E_RobotState#RS_ERROR) OR (_eState = E_RobotState#RS_RESET);
END_FUNCTION_BLOCK
